// TIA Portal V19 export
// export: Created 2026-10-15T10:10:35.7635629Z, ExportSetting WithDefaults, DisplayName Totally Integrated Automation Portal, DisplayVersion V19, DisplayName TIA Portal Openness, DisplayVersion V19, DisplayName TIA Portal Version Control Interface, DisplayVersion V19, DisplayName STEP 7 Professional, DisplayVersion V19, DisplayName STEP 7 Safety, DisplayVersion V19, DisplayName WinCC Basic/Comfort/Advanced, DisplayVersion V19, DisplayName WinCC Unified, DisplayVersion V19
FUNCTION "ROLL_PB10" : Void   // FC20, SCL
{ S7_Optimized_Access := 'TRUE' }
VERSION : 0.1
// stored: AutoNumber true, IsIECCheckEnabled false, SetENOAutomatically false, UDAEnableTagReadback false
   VAR_TEMP
      r : Bool;
      a1 : Word;
      a2 : Word;
      activeDataBlock : Int;
      comparisonResults : Array[0..0] of Bool;
   END_VAR
BEGIN

   #r := FALSE;
   #a1 := W#16#0000;
   #a2 := W#16#0000;
   #activeDataBlock := 0;
   // PB10, STEP 5 network 1
   #r := (((NOT "ROLL_State".M[110, 0]) AND (NOT "ROLL_State".M[110, 1]) AND (NOT "ROLL_State".M[110, 2]) AND (NOT "ROLL_State".M[110, 3]) AND "ROLL_State".M[40, 1]) OR ((NOT "ROLL_State".M[110, 1]) AND (NOT "ROLL_State".M[110, 2]) AND (NOT "ROLL_State".M[110, 3]) AND "ROLL_State".M[41, 2]) OR ((NOT "ROLL_State".M[110, 2]) AND (NOT "ROLL_State".M[110, 3]) AND "ROLL_State".M[42, 6]) OR ((NOT "ROLL_State".M[110, 3]) AND "ROLL_State".M[44, 2]) OR "ROLL_State".M[45, 7]);
   "ROLL_State".M[240, 0] := #r;
   // PB10, STEP 5 network 2
   #r := ((NOT "ROLL_IO".Input[119, 6]) AND "ROLL_IO".Input[12, 5] AND "ROLL_IO".Input[12, 7] AND "ROLL_State".M[110, 4] AND "ROLL_State".M[240, 0] AND "ROLL_State".M[35, 2]);
   IF #r THEN
       "ROLL_State".M[46, 2] := TRUE;
   END_IF;
   #r := ("ROLL_State".M[32, 2] OR "ROLL_State".M[46, 3]);
   IF #r THEN
       "ROLL_State".M[46, 2] := FALSE;
   END_IF;
   // PB10, STEP 5 network 3
   #r := ("ROLL_IO".Input[11, 6] AND "ROLL_IO".Input[119, 6] AND "ROLL_State".M[35, 2] AND "ROLL_State".M[46, 2]);
   IF #r THEN
       "ROLL_State".M[46, 3] := TRUE;
   END_IF;
   #r := ("ROLL_State".M[32, 2] OR "ROLL_State".M[46, 4]);
   IF #r THEN
       "ROLL_State".M[46, 3] := FALSE;
   END_IF;
   // PB10, STEP 5 network 4
   #r := ((NOT "ROLL_IO".Input[12, 1]) AND "ROLL_IO".Input[12, 5] AND "ROLL_State".M[35, 2] AND "ROLL_State".M[46, 3]);
   IF #r THEN
       "ROLL_State".M[46, 4] := TRUE;
   END_IF;
   #r := ("ROLL_State".M[32, 2] OR "ROLL_State".M[46, 5]);
   IF #r THEN
       "ROLL_State".M[46, 4] := FALSE;
   END_IF;
   // PB10, STEP 5 network 5
   #r := ("ROLL_IO".Input[12, 1] AND "ROLL_IO".Input[12, 7] AND "ROLL_State".M[35, 2] AND "ROLL_State".M[46, 4]);
   IF #r THEN
       "ROLL_State".M[46, 5] := TRUE;
   END_IF;
   #r := ("ROLL_State".M[32, 2] OR "ROLL_State".M[46, 6]);
   IF #r THEN
       "ROLL_State".M[46, 5] := FALSE;
   END_IF;
   // PB10, STEP 5 network 6
   #r := ("ROLL_State".M[35, 2] AND "ROLL_State".M[46, 5] AND "ROLL_State".S5Timers[1].Q);
   IF #r THEN
       "ROLL_State".M[46, 6] := TRUE;
   END_IF;
   #r := ("ROLL_State".M[32, 2] OR "ROLL_State".M[46, 7]);
   IF #r THEN
       "ROLL_State".M[46, 6] := FALSE;
   END_IF;
   // PB10, STEP 5 network 7
   #r := ("ROLL_State".M[35, 2] AND "ROLL_State".M[46, 6]);
   IF #r THEN
       "ROLL_State".M[46, 7] := TRUE;
   END_IF;
   #r := ("ROLL_State".M[32, 2] OR "ROLL_State".M[47, 0]);
   IF #r THEN
       "ROLL_State".M[46, 7] := FALSE;
   END_IF;
   // PB10, STEP 5 network 8
   #r := ((NOT "ROLL_IO".Input[12, 5]) AND "ROLL_State".M[35, 2] AND "ROLL_State".M[46, 7]);
   IF #r THEN
       "ROLL_State".M[47, 0] := TRUE;
   END_IF;
   #r := ("ROLL_State".M[32, 2] OR "ROLL_State".M[47, 1]);
   IF #r THEN
       "ROLL_State".M[47, 0] := FALSE;
   END_IF;
   // PB10, STEP 5 network 9
   #r := ("ROLL_IO".Input[12, 5] AND "ROLL_IO".Input[12, 7] AND "ROLL_State".M[35, 2] AND "ROLL_State".M[47, 0]);
   IF #r THEN
       "ROLL_State".M[47, 1] := TRUE;
   END_IF;
   #r := ("ROLL_State".M[32, 2] OR "ROLL_State".M[47, 2]);
   IF #r THEN
       "ROLL_State".M[47, 1] := FALSE;
   END_IF;
   // PB10, STEP 5 network 10
   #r := ("ROLL_State".M[35, 2] AND "ROLL_State".M[47, 1] AND "ROLL_State".S5Timers[2].Q);
   IF #r THEN
       "ROLL_State".M[47, 2] := TRUE;
   END_IF;
   #r := ("ROLL_State".M[32, 2] OR "ROLL_State".M[47, 3] OR "ROLL_State".M[47, 6]);
   IF #r THEN
       "ROLL_State".M[47, 2] := FALSE;
   END_IF;
   // PB10, STEP 5 network 11
   #r := ((NOT "ROLL_State".M[110, 5]) AND (NOT "ROLL_State".M[110, 6]) AND "ROLL_State".M[35, 2] AND "ROLL_State".M[47, 2]);
   IF #r THEN
       "ROLL_State".M[47, 3] := TRUE;
   END_IF;
   #r := ("ROLL_State".M[32, 2] OR "ROLL_State".M[47, 4]);
   IF #r THEN
       "ROLL_State".M[47, 3] := FALSE;
   END_IF;
   // PB10, STEP 5 network 12
   #r := ("ROLL_IO".Input[13, 3] AND "ROLL_State".M[35, 2] AND "ROLL_State".M[47, 3] AND "ROLL_State".M[63, 1]);
   IF #r THEN
       "ROLL_State".M[47, 4] := TRUE;
   END_IF;
   #r := ("ROLL_State".M[32, 2] OR "ROLL_State".M[50, 6] OR "ROLL_State".M[52, 0]);
   IF #r THEN
       "ROLL_State".M[47, 4] := FALSE;
   END_IF;
   // PB10, STEP 5 network 13
   #r := (((NOT "ROLL_State".M[110, 0]) AND (NOT "ROLL_State".M[110, 1]) AND (NOT "ROLL_State".M[110, 2]) AND (NOT "ROLL_State".M[110, 3]) AND (NOT "ROLL_State".M[110, 4]) AND "ROLL_State".M[40, 1]) OR ((NOT "ROLL_State".M[110, 1]) AND (NOT "ROLL_State".M[110, 2]) AND (NOT "ROLL_State".M[110, 3]) AND (NOT "ROLL_State".M[110, 4]) AND "ROLL_State".M[41, 2]) OR ((NOT "ROLL_State".M[110, 2]) AND (NOT "ROLL_State".M[110, 3]) AND (NOT "ROLL_State".M[110, 4]) AND "ROLL_State".M[42, 6]) OR ((NOT "ROLL_State".M[110, 3]) AND (NOT "ROLL_State".M[110, 4]) AND "ROLL_State".M[44, 2]) OR ((NOT "ROLL_State".M[110, 4]) AND "ROLL_State".M[45, 7]) OR "ROLL_State".M[47, 2]);
   "ROLL_State".M[240, 0] := #r;
   // PB10, STEP 5 network 14
   #r := ((NOT "ROLL_IO".Input[119, 7]) AND "ROLL_IO".Input[12, 5] AND "ROLL_IO".Input[12, 7] AND "ROLL_State".M[110, 5] AND "ROLL_State".M[240, 0] AND "ROLL_State".M[35, 2]);
   IF #r THEN
       "ROLL_State".M[47, 6] := TRUE;
   END_IF;
   #r := ("ROLL_State".M[32, 2] OR "ROLL_State".M[47, 7]);
   IF #r THEN
       "ROLL_State".M[47, 6] := FALSE;
   END_IF;
   // PB10, STEP 5 network 15
   #r := ("ROLL_IO".Input[11, 6] AND "ROLL_IO".Input[119, 7] AND "ROLL_State".M[35, 2] AND "ROLL_State".M[47, 6]);
   IF #r THEN
       "ROLL_State".M[47, 7] := TRUE;
   END_IF;
   #r := ("ROLL_State".M[32, 2] OR "ROLL_State".M[48, 0]);
   IF #r THEN
       "ROLL_State".M[47, 7] := FALSE;
   END_IF;
   // PB10, STEP 5 network 16
   #r := ((NOT "ROLL_IO".Input[12, 1]) AND "ROLL_IO".Input[12, 5] AND "ROLL_State".M[35, 2] AND "ROLL_State".M[47, 7]);
   IF #r THEN
       "ROLL_State".M[48, 0] := TRUE;
   END_IF;
   #r := ("ROLL_State".M[32, 2] OR "ROLL_State".M[48, 1]);
   IF #r THEN
       "ROLL_State".M[48, 0] := FALSE;
   END_IF;
   // PB10, STEP 5 network 17
   #r := ("ROLL_IO".Input[12, 1] AND "ROLL_IO".Input[12, 7] AND "ROLL_State".M[35, 2] AND "ROLL_State".M[48, 0]);
   IF #r THEN
       "ROLL_State".M[48, 1] := TRUE;
   END_IF;
   #r := ("ROLL_State".M[32, 2] OR "ROLL_State".M[48, 2]);
   IF #r THEN
       "ROLL_State".M[48, 1] := FALSE;
   END_IF;
   // PB10, STEP 5 network 18
   #r := ("ROLL_State".M[35, 2] AND "ROLL_State".M[48, 1] AND "ROLL_State".S5Timers[1].Q);
   IF #r THEN
       "ROLL_State".M[48, 2] := TRUE;
   END_IF;
   #r := ("ROLL_State".M[32, 2] OR "ROLL_State".M[48, 3]);
   IF #r THEN
       "ROLL_State".M[48, 2] := FALSE;
   END_IF;
   // PB10, STEP 5 network 19
   #r := ("ROLL_State".M[35, 2] AND "ROLL_State".M[48, 2]);
   IF #r THEN
       "ROLL_State".M[48, 3] := TRUE;
   END_IF;
   #r := ("ROLL_State".M[32, 2] OR "ROLL_State".M[48, 4]);
   IF #r THEN
       "ROLL_State".M[48, 3] := FALSE;
   END_IF;
   // PB10, STEP 5 network 20
   #r := ((NOT "ROLL_IO".Input[12, 5]) AND "ROLL_State".M[35, 2] AND "ROLL_State".M[48, 3]);
   IF #r THEN
       "ROLL_State".M[48, 4] := TRUE;
   END_IF;
   #r := ("ROLL_State".M[32, 2] OR "ROLL_State".M[48, 5]);
   IF #r THEN
       "ROLL_State".M[48, 4] := FALSE;
   END_IF;
   // PB10, STEP 5 network 21
   #r := ("ROLL_IO".Input[12, 5] AND "ROLL_IO".Input[12, 7] AND "ROLL_State".M[35, 2] AND "ROLL_State".M[48, 4]);
   IF #r THEN
       "ROLL_State".M[48, 5] := TRUE;
   END_IF;
   #r := ("ROLL_State".M[32, 2] OR "ROLL_State".M[48, 6]);
   IF #r THEN
       "ROLL_State".M[48, 5] := FALSE;
   END_IF;
   // PB10, STEP 5 network 22
   #r := ("ROLL_State".M[35, 2] AND "ROLL_State".M[48, 5] AND "ROLL_State".S5Timers[2].Q);
   IF #r THEN
       "ROLL_State".M[48, 6] := TRUE;
   END_IF;
   #r := ("ROLL_State".M[32, 2] OR "ROLL_State".M[48, 7] OR "ROLL_State".M[49, 2]);
   IF #r THEN
       "ROLL_State".M[48, 6] := FALSE;
   END_IF;
   // PB10, STEP 5 network 23
   #r := ((NOT "ROLL_State".M[110, 6]) AND "ROLL_State".M[35, 2] AND "ROLL_State".M[48, 6]);
   IF #r THEN
       "ROLL_State".M[48, 7] := TRUE;
   END_IF;
   #r := ("ROLL_State".M[32, 2] OR "ROLL_State".M[49, 0]);
   IF #r THEN
       "ROLL_State".M[48, 7] := FALSE;
   END_IF;
   // PB10, STEP 5 network 24
   #r := ("ROLL_IO".Input[13, 3] AND "ROLL_State".M[35, 2] AND "ROLL_State".M[48, 7] AND "ROLL_State".M[63, 1]);
   IF #r THEN
       "ROLL_State".M[49, 0] := TRUE;
   END_IF;
   #r := ("ROLL_State".M[32, 2] OR "ROLL_State".M[50, 6] OR "ROLL_State".M[52, 0]);
   IF #r THEN
       "ROLL_State".M[49, 0] := FALSE;
   END_IF;
   // PB10, STEP 5 network 25
   #r := (((NOT "ROLL_State".M[110, 0]) AND (NOT "ROLL_State".M[110, 1]) AND (NOT "ROLL_State".M[110, 2]) AND (NOT "ROLL_State".M[110, 3]) AND (NOT "ROLL_State".M[110, 4]) AND (NOT "ROLL_State".M[110, 5]) AND "ROLL_State".M[40, 1]) OR ((NOT "ROLL_State".M[110, 1]) AND (NOT "ROLL_State".M[110, 2]) AND (NOT "ROLL_State".M[110, 3]) AND (NOT "ROLL_State".M[110, 4]) AND (NOT "ROLL_State".M[110, 5]) AND "ROLL_State".M[41, 2]) OR ((NOT "ROLL_State".M[110, 2]) AND (NOT "ROLL_State".M[110, 3]) AND (NOT "ROLL_State".M[110, 4]) AND (NOT "ROLL_State".M[110, 5]) AND "ROLL_State".M[42, 6]) OR ((NOT "ROLL_State".M[110, 3]) AND (NOT "ROLL_State".M[110, 4]) AND (NOT "ROLL_State".M[110, 5]) AND "ROLL_State".M[44, 2]) OR ((NOT "ROLL_State".M[110, 4]) AND (NOT "ROLL_State".M[110, 5]) AND "ROLL_State".M[45, 7]) OR ((NOT "ROLL_State".M[110, 5]) AND "ROLL_State".M[47, 2]) OR "ROLL_State".M[48, 6]);
   "ROLL_State".M[240, 0] := #r;
   // PB10, STEP 5 network 26
   #r := ((NOT "ROLL_IO".Input[120, 0]) AND "ROLL_IO".Input[12, 5] AND "ROLL_IO".Input[12, 7] AND "ROLL_State".M[110, 6] AND "ROLL_State".M[240, 0] AND "ROLL_State".M[35, 2]);
   IF #r THEN
       "ROLL_State".M[49, 2] := TRUE;
   END_IF;
   #r := ("ROLL_State".M[32, 2] OR "ROLL_State".M[49, 3]);
   IF #r THEN
       "ROLL_State".M[49, 2] := FALSE;
   END_IF;
   // PB10, STEP 5 network 27
   #r := ("ROLL_IO".Input[11, 6] AND "ROLL_IO".Input[120, 0] AND "ROLL_State".M[35, 2] AND "ROLL_State".M[49, 2]);
   IF #r THEN
       "ROLL_State".M[49, 3] := TRUE;
   END_IF;
   #r := ("ROLL_State".M[32, 2] OR "ROLL_State".M[49, 4]);
   IF #r THEN
       "ROLL_State".M[49, 3] := FALSE;
   END_IF;
   // PB10, STEP 5 network 28
   #r := ((NOT "ROLL_IO".Input[12, 1]) AND "ROLL_IO".Input[12, 5] AND "ROLL_State".M[35, 2] AND "ROLL_State".M[49, 3]);
   IF #r THEN
       "ROLL_State".M[49, 4] := TRUE;
   END_IF;
   #r := ("ROLL_State".M[32, 2] OR "ROLL_State".M[49, 5]);
   IF #r THEN
       "ROLL_State".M[49, 4] := FALSE;
   END_IF;
   // PB10, STEP 5 network 29
   #r := ("ROLL_IO".Input[12, 1] AND "ROLL_IO".Input[12, 7] AND "ROLL_State".M[35, 2] AND "ROLL_State".M[49, 4]);
   IF #r THEN
       "ROLL_State".M[49, 5] := TRUE;
   END_IF;
   #r := ("ROLL_State".M[32, 2] OR "ROLL_State".M[49, 6]);
   IF #r THEN
       "ROLL_State".M[49, 5] := FALSE;
   END_IF;
   // PB10, STEP 5 network 30
   #r := ("ROLL_State".M[35, 2] AND "ROLL_State".M[49, 5] AND "ROLL_State".S5Timers[1].Q);
   IF #r THEN
       "ROLL_State".M[49, 6] := TRUE;
   END_IF;
   #r := ("ROLL_State".M[32, 2] OR "ROLL_State".M[49, 7]);
   IF #r THEN
       "ROLL_State".M[49, 6] := FALSE;
   END_IF;
   // PB10, STEP 5 network 31
   #r := ("ROLL_State".M[35, 2] AND "ROLL_State".M[49, 6]);
   IF #r THEN
       "ROLL_State".M[49, 7] := TRUE;
   END_IF;
   #r := ("ROLL_State".M[32, 2] OR "ROLL_State".M[50, 0]);
   IF #r THEN
       "ROLL_State".M[49, 7] := FALSE;
   END_IF;
   // PB10, STEP 5 network 32
   #r := ((NOT "ROLL_IO".Input[12, 5]) AND "ROLL_State".M[35, 2] AND "ROLL_State".M[49, 7]);
   IF #r THEN
       "ROLL_State".M[50, 0] := TRUE;
   END_IF;
   #r := ("ROLL_State".M[32, 2] OR "ROLL_State".M[50, 1]);
   IF #r THEN
       "ROLL_State".M[50, 0] := FALSE;
   END_IF;
   // PB10, STEP 5 network 33
   #r := ("ROLL_IO".Input[12, 5] AND "ROLL_IO".Input[12, 7] AND "ROLL_State".M[35, 2] AND "ROLL_State".M[50, 0]);
   IF #r THEN
       "ROLL_State".M[50, 1] := TRUE;
   END_IF;
   #r := ("ROLL_State".M[32, 2] OR "ROLL_State".M[50, 2]);
   IF #r THEN
       "ROLL_State".M[50, 1] := FALSE;
   END_IF;
   // PB10, STEP 5 network 34
   #r := ("ROLL_State".M[35, 2] AND "ROLL_State".M[50, 1] AND "ROLL_State".S5Timers[2].Q);
   IF #r THEN
       "ROLL_State".M[50, 2] := TRUE;
   END_IF;
   #r := ("ROLL_State".M[32, 2] OR "ROLL_State".M[50, 3]);
   IF #r THEN
       "ROLL_State".M[50, 2] := FALSE;
   END_IF;
   // PB10, STEP 5 network 35
   #r := ("ROLL_State".M[35, 2] AND "ROLL_State".M[50, 2]);
   IF #r THEN
       "ROLL_State".M[50, 3] := TRUE;
   END_IF;
   #r := ("ROLL_State".M[32, 2] OR "ROLL_State".M[50, 4]);
   IF #r THEN
       "ROLL_State".M[50, 3] := FALSE;
   END_IF;
   // PB10, STEP 5 network 36
   #r := ("ROLL_IO".Input[13, 3] AND "ROLL_State".M[35, 2] AND "ROLL_State".M[50, 3] AND "ROLL_State".M[63, 1]);
   IF #r THEN
       "ROLL_State".M[50, 4] := TRUE;
   END_IF;
   #r := ("ROLL_State".M[32, 2] OR "ROLL_State".M[50, 6] OR "ROLL_State".M[52, 0]);
   IF #r THEN
       "ROLL_State".M[50, 4] := FALSE;
   END_IF;
   // PB10, STEP 5 network 37
   #r := (((NOT "ROLL_State".M[110, 0]) AND (NOT "ROLL_State".M[110, 1]) AND (NOT "ROLL_State".M[110, 2]) AND (NOT "ROLL_State".M[110, 3]) AND (NOT "ROLL_State".M[110, 4]) AND (NOT "ROLL_State".M[110, 5]) AND (NOT "ROLL_State".M[110, 6]) AND "ROLL_State".M[40, 1]) OR ((NOT "ROLL_State".M[110, 1]) AND (NOT "ROLL_State".M[110, 2]) AND (NOT "ROLL_State".M[110, 3]) AND (NOT "ROLL_State".M[110, 4]) AND (NOT "ROLL_State".M[110, 5]) AND (NOT "ROLL_State".M[110, 6]) AND "ROLL_State".M[41, 4]) OR ((NOT "ROLL_State".M[110, 2]) AND (NOT "ROLL_State".M[110, 3]) AND (NOT "ROLL_State".M[110, 4]) AND (NOT "ROLL_State".M[110, 5]) AND (NOT "ROLL_State".M[110, 6]) AND "ROLL_State".M[43, 0]));
   "ROLL_State".M[240, 0] := #r;
   // PB10, STEP 5 network 38
   #r := (((NOT "ROLL_State".M[110, 3]) AND (NOT "ROLL_State".M[110, 4]) AND (NOT "ROLL_State".M[110, 5]) AND (NOT "ROLL_State".M[110, 6]) AND "ROLL_State".M[44, 4]) OR ((NOT "ROLL_State".M[110, 4]) AND (NOT "ROLL_State".M[110, 5]) AND (NOT "ROLL_State".M[110, 6]) AND "ROLL_State".M[46, 1]) OR ((NOT "ROLL_State".M[110, 5]) AND (NOT "ROLL_State".M[110, 6]) AND "ROLL_State".M[47, 4]) OR ((NOT "ROLL_State".M[110, 6]) AND "ROLL_State".M[49, 0]) OR "ROLL_State".M[50, 4]);
   "ROLL_State".M[240, 1] := #r;
   // PB10, STEP 5 network 39
   #r := ((NOT "ROLL_IO".Input[120, 1]) AND ("ROLL_State".M[240, 0] OR "ROLL_State".M[240, 1]) AND "ROLL_IO".Input[12, 5] AND "ROLL_IO".Input[12, 7] AND "ROLL_State".M[110, 7] AND "ROLL_State".M[35, 2] AND "ROLL_State".M[63, 1]);
   IF #r THEN
       "ROLL_State".M[50, 6] := TRUE;
   END_IF;
   #r := ("ROLL_State".M[32, 2] OR "ROLL_State".M[50, 7]);
   IF #r THEN
       "ROLL_State".M[50, 6] := FALSE;
   END_IF;
   // PB10, STEP 5 network 40
   #r := ("ROLL_IO".Input[11, 6] AND "ROLL_IO".Input[120, 1] AND "ROLL_State".M[35, 2] AND "ROLL_State".M[50, 6]);
   IF #r THEN
       "ROLL_State".M[50, 7] := TRUE;
   END_IF;
   #r := ("ROLL_State".M[32, 2] OR "ROLL_State".M[51, 0]);
   IF #r THEN
       "ROLL_State".M[50, 7] := FALSE;
   END_IF;
   // PB10, STEP 5 network 41
   #r := ((NOT "ROLL_IO".Input[12, 1]) AND "ROLL_IO".Input[12, 5] AND "ROLL_State".M[35, 2] AND "ROLL_State".M[50, 7]);
   IF #r THEN
       "ROLL_State".M[51, 0] := TRUE;
   END_IF;
   #r := ("ROLL_State".M[32, 2] OR "ROLL_State".M[51, 1]);
   IF #r THEN
       "ROLL_State".M[51, 0] := FALSE;
   END_IF;
   // PB10, STEP 5 network 42
   #r := ("ROLL_State".M[35, 2] AND "ROLL_State".M[51, 0] AND "ROLL_State".M[80, 6]);
   IF #r THEN
       "ROLL_State".M[51, 1] := TRUE;
   END_IF;
   #r := ("ROLL_State".M[32, 2] OR "ROLL_State".M[51, 2]);
   IF #r THEN
       "ROLL_State".M[51, 1] := FALSE;
   END_IF;
   // PB10, STEP 5 network 43
   #r := ("ROLL_State".M[35, 2] AND "ROLL_State".M[51, 1] AND "ROLL_State".S5Timers[1].Q);
   IF #r THEN
       "ROLL_State".M[51, 2] := TRUE;
   END_IF;
   #r := ("ROLL_State".M[32, 2] OR "ROLL_State".M[51, 3]);
   IF #r THEN
       "ROLL_State".M[51, 2] := FALSE;
   END_IF;
   // PB10, STEP 5 network 44
   #r := ((NOT "ROLL_IO".Input[12, 5]) AND "ROLL_State".M[35, 2] AND "ROLL_State".M[51, 2]);
   IF #r THEN
       "ROLL_State".M[51, 3] := TRUE;
   END_IF;
   #r := ("ROLL_State".M[32, 2] OR "ROLL_State".M[51, 4]);
   IF #r THEN
       "ROLL_State".M[51, 3] := FALSE;
   END_IF;
   // PB10, STEP 5 network 45
   #r := ("ROLL_IO".Input[12, 5] AND "ROLL_IO".Input[12, 7] AND "ROLL_State".M[35, 2] AND "ROLL_State".M[51, 3]);
   IF #r THEN
       "ROLL_State".M[51, 4] := TRUE;
   END_IF;
   #r := ("ROLL_State".M[32, 2] OR "ROLL_State".M[51, 5]);
   IF #r THEN
       "ROLL_State".M[51, 4] := FALSE;
   END_IF;
   // PB10, STEP 5 network 46
   #r := ("ROLL_State".M[35, 2] AND "ROLL_State".M[51, 4]);
   IF #r THEN
       "ROLL_State".M[51, 5] := TRUE;
   END_IF;
   #r := ("ROLL_State".M[32, 2] OR "ROLL_State".M[51, 6]);
   IF #r THEN
       "ROLL_State".M[51, 5] := FALSE;
   END_IF;
   // PB10, STEP 5 network 47
   #r := ("ROLL_IO".Input[13, 3] AND "ROLL_State".M[35, 2] AND "ROLL_State".M[51, 5] AND "ROLL_State".M[63, 1]);
   IF #r THEN
       "ROLL_State".M[51, 6] := TRUE;
   END_IF;
   #r := ("ROLL_State".M[32, 2] OR "ROLL_State".M[52, 0]);
   IF #r THEN
       "ROLL_State".M[51, 6] := FALSE;
   END_IF;
   // PB10, STEP 5 network 48
   #r := (((NOT "ROLL_State".M[110, 1]) AND (NOT "ROLL_State".M[110, 2]) AND (NOT "ROLL_State".M[110, 3]) AND (NOT "ROLL_State".M[110, 4]) AND (NOT "ROLL_State".M[110, 5]) AND (NOT "ROLL_State".M[110, 6]) AND (NOT "ROLL_State".M[110, 7]) AND "ROLL_State".M[41, 4]) OR ((NOT "ROLL_State".M[110, 2]) AND (NOT "ROLL_State".M[110, 3]) AND (NOT "ROLL_State".M[110, 4]) AND (NOT "ROLL_State".M[110, 5]) AND (NOT "ROLL_State".M[110, 6]) AND (NOT "ROLL_State".M[110, 7]) AND "ROLL_State".M[43, 0]));
   "ROLL_State".M[240, 0] := #r;
   // PB10, STEP 5 network 49
   #r := (((NOT "ROLL_State".M[110, 3]) AND (NOT "ROLL_State".M[110, 4]) AND (NOT "ROLL_State".M[110, 5]) AND (NOT "ROLL_State".M[110, 6]) AND (NOT "ROLL_State".M[110, 7]) AND "ROLL_State".M[44, 4]) OR ((NOT "ROLL_State".M[110, 4]) AND (NOT "ROLL_State".M[110, 5]) AND (NOT "ROLL_State".M[110, 6]) AND (NOT "ROLL_State".M[110, 7]) AND "ROLL_State".M[46, 1]) OR ((NOT "ROLL_State".M[110, 5]) AND (NOT "ROLL_State".M[110, 6]) AND (NOT "ROLL_State".M[110, 7]) AND "ROLL_State".M[47, 4]) OR ((NOT "ROLL_State".M[110, 6]) AND (NOT "ROLL_State".M[110, 7]) AND "ROLL_State".M[49, 0]) OR ((NOT "ROLL_State".M[110, 7]) AND "ROLL_State".M[50, 4]) OR "ROLL_State".M[51, 6]);
   "ROLL_State".M[240, 1] := #r;
   // PB10, STEP 5 network 50
   #r := ((NOT "ROLL_IO".Input[11, 0]) AND ("ROLL_State".M[240, 0] OR "ROLL_State".M[240, 1]) AND "ROLL_IO".Input[12, 5] AND "ROLL_IO".Input[12, 7] AND "ROLL_IO".Input[13, 3] AND "ROLL_State".M[35, 2] AND "ROLL_State".M[63, 1]);
   IF #r THEN
       "ROLL_State".M[52, 0] := TRUE;
   END_IF;
   #r := ("ROLL_State".M[32, 2] OR "ROLL_State".M[52, 1]);
   IF #r THEN
       "ROLL_State".M[52, 0] := FALSE;
   END_IF;
   // PB10, STEP 5 network 51
   #r := ("ROLL_IO".Input[11, 0] AND "ROLL_IO".Input[11, 6] AND "ROLL_State".M[35, 2] AND "ROLL_State".M[52, 0]);
   IF #r THEN
       "ROLL_State".M[52, 1] := TRUE;
   END_IF;
   #r := ("ROLL_State".M[32, 2] OR "ROLL_State".M[52, 2]);
   IF #r THEN
       "ROLL_State".M[52, 1] := FALSE;
   END_IF;
   // PB10, STEP 5 network 52
   #r := ((NOT "ROLL_IO".Input[12, 1]) AND (("ROLL_IO".Input[124, 2] AND "ROLL_IO".Input[124, 5]) OR "ROLL_State".M[0, 4]) AND "ROLL_IO".Input[12, 5] AND "ROLL_State".M[35, 2] AND "ROLL_State".M[52, 1]);
   IF #r THEN
       "ROLL_State".M[52, 2] := TRUE;
   END_IF;
   #r := ("ROLL_State".M[32, 2] OR "ROLL_State".M[52, 3]);
   IF #r THEN
       "ROLL_State".M[52, 2] := FALSE;
   END_IF;
   // PB10, STEP 5 network 53
   #r := ("ROLL_IO".Input[12, 1] AND "ROLL_IO".Input[12, 7] AND "ROLL_State".M[35, 2] AND "ROLL_State".M[52, 2]);
   IF #r THEN
       "ROLL_State".M[52, 3] := TRUE;
   END_IF;
   #r := ("ROLL_State".M[32, 2] OR "ROLL_State".M[53, 0] OR "ROLL_State".M[53, 6]);
   IF #r THEN
       "ROLL_State".M[52, 3] := FALSE;
   END_IF;
   // PB10, STEP 5 network 54
   #r := ((NOT "ROLL_IO".Output[113, 3]) AND (NOT "ROLL_IO".Input[123, 5]) AND (NOT "ROLL_IO".Input[123, 6]) AND (NOT "ROLL_IO".Input[124, 1]) AND (NOT "ROLL_State".M[70, 3]) AND "ROLL_IO".Output[113, 2] AND "ROLL_IO".Input[124, 2] AND "ROLL_State".M[0, 3] AND "ROLL_State".M[35, 2] AND "ROLL_State".M[52, 3]);
   IF #r THEN
       "ROLL_State".M[53, 0] := TRUE;
   END_IF;
   #r := ("ROLL_State".M[32, 2] OR "ROLL_State".M[53, 1]);
   IF #r THEN
       "ROLL_State".M[53, 0] := FALSE;
   END_IF;
   // PB10, STEP 5 network 55
   #r := ((NOT "ROLL_IO".Input[124, 2]) AND "ROLL_IO".Input[124, 1] AND "ROLL_State".M[35, 2] AND "ROLL_State".M[53, 0]);
   IF #r THEN
       "ROLL_State".M[53, 1] := TRUE;
   END_IF;
   #r := ("ROLL_State".M[32, 2] OR "ROLL_State".M[53, 2]);
   IF #r THEN
       "ROLL_State".M[53, 1] := FALSE;
   END_IF;
   // PB10, STEP 5 network 56
   #r := ((NOT "ROLL_IO".Input[124, 4]) AND "ROLL_IO".Input[124, 5] AND "ROLL_State".M[35, 2] AND "ROLL_State".M[53, 1]);
   IF #r THEN
       "ROLL_State".M[53, 2] := TRUE;
   END_IF;
   #r := ("ROLL_State".M[32, 2] OR "ROLL_State".M[53, 3]);
   IF #r THEN
       "ROLL_State".M[53, 2] := FALSE;
   END_IF;
   // PB10, STEP 5 network 57
   #r := ((NOT "ROLL_IO".Input[124, 5]) AND "ROLL_IO".Input[124, 4] AND "ROLL_State".M[35, 2] AND "ROLL_State".M[53, 2]);
   IF #r THEN
       "ROLL_State".M[53, 3] := TRUE;
   END_IF;
   #r := ("ROLL_State".M[32, 2] OR "ROLL_State".M[53, 4]);
   IF #r THEN
       "ROLL_State".M[53, 3] := FALSE;
   END_IF;
   // PB10, STEP 5 network 58
   #r := ((NOT "ROLL_State".M[53, 2]) AND "ROLL_State".M[35, 2] AND "ROLL_State".M[53, 3]);
   IF #r THEN
       "ROLL_State".M[53, 4] := TRUE;
   END_IF;
   #r := ("ROLL_State".M[32, 2] OR "ROLL_State".M[53, 5]);
   IF #r THEN
       "ROLL_State".M[53, 4] := FALSE;
   END_IF;
   // PB10, STEP 5 network 59
   #r := ((NOT "ROLL_IO".Input[123, 5]) AND (NOT "ROLL_IO".Input[123, 6]) AND (NOT "ROLL_State".M[70, 3]) AND "ROLL_State".M[35, 2] AND "ROLL_State".M[53, 4]);
   IF #r THEN
       "ROLL_State".M[53, 5] := TRUE;
   END_IF;
   #r := ("ROLL_State".M[32, 2] OR "ROLL_State".M[53, 6]);
   IF #r THEN
       "ROLL_State".M[53, 5] := FALSE;
   END_IF;
   // PB10, STEP 5 network 60
   #r := (("ROLL_State".M[52, 3] OR "ROLL_State".M[53, 5]) AND "ROLL_State".M[35, 2]);
   IF #r THEN
       "ROLL_State".M[53, 6] := TRUE;
   END_IF;
   #r := ("ROLL_State".M[32, 2] OR "ROLL_State".M[37, 0]);
   IF #r THEN
       "ROLL_State".M[53, 6] := FALSE;
   END_IF;
   // PB10, STEP 5 network 61
   RETURN;
END_FUNCTION
